(* IEC 61131-3 sources: Test-Git_ESME26/TestProgettoESME_26.fbsproj/PacDriveLib Migration/Motion/Homing/PDL_FB_SetTrackingDeviation.fb.st^, 4 files *)

(* ---- ifDrive2.prop.st ---- *)
PROPERTY PUBLIC ifDrive2 : DDI.IF_Drive2;

__SETTERDECLARATION__
VAR
END_VAR
__SETTERIMPLEMENTATION__
ifDrive2_loc := ifDrive2;

(* ---- lrCurrentTrackDevLim.prop.st ---- *)
PROPERTY PUBLIC lrCurrentTrackDevLim : LREAL
__GETTERDECLARATION__
VAR
END_VAR
__GETTERIMPLEMENTATION__
lrCurrentTrackDevLim := lrCurrentTrackingDeviationLimit;
__SETTERDECLARATION__
VAR
END_VAR
__SETTERIMPLEMENTATION__

(* ---- lrOldTrackDevLim.prop.st ---- *)
PROPERTY PUBLIC lrOldTrackDevLim : LREAL
__SETTERDECLARATION__
VAR
END_VAR
__SETTERIMPLEMENTATION__

__GETTERDECLARATION__
VAR
END_VAR
__GETTERIMPLEMENTATION__
lrOldTrackDevLim := lrOldTrackingDeviationLimit;

(* ---- xDone.prop.st ---- *)
PROPERTY xDone : BOOL
__GETTERDECLARATION__
VAR
END_VAR
__GETTERIMPLEMENTATION__
xDone := xDone_loc;
__SETTERDECLARATION__
VAR
END_VAR
__SETTERIMPLEMENTATION__
xDone_loc := xDone;
